FUNCTION_BLOCK FB_ActuatorModulating EXTENDS FB_Device
(*
	Continuous-position actuator: control valve, damper, any 0-100 % analog-positioned device.
	0 % = closed, 100 % = open. The output ramps to the setpoint at cfg.rampRate and is
	scaled to raw counts for an analog output terminal.
	
	Interlocks: losing them moves the actuator to cfg.safePosition. Permissives are required
	to move away from the safe position.
	
	Feedback: position comes from positionFdbk (FB_AnalogInput). In simulation, or with
	cfg.noFdbk, the position follows the output at the speed set by cfg.strokeTime.
	Simulation holds the physical output at 0.
*)
VAR_INPUT
	{attribute 'OPC.UA.DA' := '1'}
	{attribute 'OPC.UA.DA.StructuredType' := '1'}
	cfg					: ST_ActuatorModulatingConfiguration; //configuration
	
	{attribute 'OPC.UA.DA' := '1'}
	ocmd				: E_ActuatorModulatingCommand; //operator command
	{attribute 'OPC.UA.DA' := '1'}
	opPosition			: LREAL; //operator target position in %, used with ocmd Position
	
	func				: ST_ActuatorModulatingFunctions; //functions
	
	(* Interlocks/Permissives
	----------------------------------------------------------------------------------------------------*)
	{attribute 'OPC.UA.DA' := '1'}
	{attribute 'OPC.UA.DA.Access' := '1'}
	intlk				: FB_Permissive; //losing these moves the actuator to safePosition
	{attribute 'OPC.UA.DA' := '1'}
	{attribute 'OPC.UA.DA.Access' := '1'}
	perm				: FB_Permissive; //required to move away from safePosition
	
	(* External inputs
	----------------------------------------------------------------------------------------------------*)
	{attribute 'OPC.UA.DA' := '1'}
	{attribute 'OPC.UA.DA.Access' := '1'}
	positionFdbk		: FB_AnalogInput; //position feedback, link positionFdbk.inpRaw
END_VAR
VAR_OUTPUT
	outRaw		AT %Q*	: INT; //analog output to the actuator, link to the terminal's Value
	
	{attribute 'OPC.UA.DA' := '1'}
	{attribute 'OPC.UA.DA.Access' := '1'}
	{attribute 'OPC.UA.DA.StructuredType' := '1'}
	sts					: ST_ActuatorModulatingStatus;
	
	{attribute 'OPC.UA.DA' := '1'}
	{attribute 'OPC.UA.DA.Access' := '1'}
	{attribute 'OPC.UA.DA.StructuredType' := '1'}
	fault				: ST_ActuatorModulatingFault;
END_VAR
VAR
	//Command processing
	pcmd				: E_ActuatorModulatingCommand; //program command
	pPosition			: LREAL; //program target position in %, used with pcmd Position
	pcmdLast			: E_ActuatorModulatingCommand;
	ocmdLast			: E_ActuatorModulatingCommand;
	cmdReceived			: E_ActuatorModulatingCommand; //command accepted this scan
	targetReceived		: LREAL; //target position that came with cmdReceived
	funcTarget			: LREAL; //target of the running ToPosition function
	
	//state variables for tracking
	stateLastScan		: E_ActuatorModulatingState; //state on last scan
	simPosition			: LREAL; //simulated position in %
	
	//Oneshot triggers
	rtNewState			: BOOL; //just entered new state
	
	//Timers
	deltaTime			: FB_DeltaTime; //scan time for ramp and simulation
	positioningTimer	: TON; //time spent positioning
	
	resetFault			: BOOL;
END_VAR

SUPER^();

Device();
StatusIn();
ProcessInputs();
ProcessCommands();
Functions();
StateMachine();
HandleFaults();
ControlOutputs();
StatusOut();

METHOD PUBLIC Close
pcmd := E_ActuatorModulatingCommand.Close;
END_METHOD

METHOD PROTECTED ControlOutputs //Set physical outputs
IF sts.sim THEN //do not command outputs when simulated
	outRaw := 0;
ELSE
	outRaw := LREAL_TO_INT(F_ScaleLinear(value := sts.commandPosition, inMin := 0, inMax := 100,
										outMin := cfg.outRawAtClosed, outMax := cfg.outRawAtOpen, clamp := TRUE));
END_IF
END_METHOD

METHOD PROTECTED Device //map cfg to FB_Device and FB_Device to sts
// to FB device
opTimeout  			 := cfg.opTimeout;
opTimeoutEnable 	 := cfg.opTimeoutEnable;
opActivity 			 := ocmd <> E_ActuatorModulatingCommand.None;

// from FB device
sts.mode	   		 := mode;
sts.modeAuto   		 := sts.mode = E_SystemMode.Auto;
sts.modeManual 		 := sts.mode = E_SystemMode.Manual;
sts.manualOvrde		 := ctrl.manualOvrde;
sts.bypass 	   		 := ctrl.bypass;
sts.sim		   		 := ctrl.sim;
sts.parentConfigured := parentConfigured;
END_METHOD

METHOD PROTECTED Functions
VAR
	i : INT;
END_VAR
func.ToPosition(hmiTextStatic := CONCAT(cfg.actuatorId, ' to position'), timeoutPT := cfg.failTimePositioning);
func.ToPosition.permComplete.cfg.condText[0] := CONCAT(cfg.actuatorId, ' at position');
IF func.ToPosition.entry THEN
	funcTarget := sts.setpoint; // no Position parameter = stay where it is
	FOR i := GVL_Lib_SequencerConstants.MIN_PARAMETERS TO GVL_Lib_SequencerConstants.MAX_PARAMETERS DO
		IF func.ToPosition.arrParam[i].typeEnum = E_ActuatorModulatingFunctionParam.Position THEN
			funcTarget := func.ToPosition.arrParam[i].value;
		END_IF
	END_FOR
	SetPosition(funcTarget);
END_IF
IF func.ToPosition.running THEN
	func.ToPosition.permComplete.perm.0 := sts.atPosition AND ABS(sts.setpoint - LIMIT(cfg.minPosition, funcTarget, cfg.maxPosition)) < 0.001;
	IF NOT func.ToPosition.permComplete.perm.0 AND ABS(sts.setpoint - funcTarget) >= 0.001 AND NOT fault.active THEN
		SetPosition(funcTarget); // continue calling if didn't work at first
	END_IF
	func.ToPosition.inpError := fault.active;
	func.ToPosition.inpErrorText := fault.text;
END_IF


func.Open(hmiTextStatic := CONCAT(cfg.actuatorId, ' open'), timeoutPT := cfg.failTimePositioning);
func.Open.permComplete.cfg.condText[0] := CONCAT(cfg.actuatorId, ' open');
func.Open.permComplete.perm.0 := sts.atPosition AND sts.setpoint = cfg.maxPosition;
IF func.Open.entry OR (func.Open.running AND sts.setpoint <> cfg.maxPosition AND NOT fault.active) THEN
	Open();
END_IF
IF func.Open.running THEN
	func.Open.inpError := fault.active;
	func.Open.inpErrorText := fault.text;
END_IF


func.Close(hmiTextStatic := CONCAT(cfg.actuatorId, ' close'), timeoutPT := cfg.failTimePositioning);
func.Close.permComplete.cfg.condText[0] := CONCAT(cfg.actuatorId, ' closed');
func.Close.permComplete.perm.0 := sts.atPosition AND sts.setpoint = cfg.minPosition;
IF func.Close.entry OR (func.Close.running AND sts.setpoint <> cfg.minPosition AND NOT fault.active) THEN
	Close();
END_IF
IF func.Close.running THEN
	func.Close.inpError := fault.active;
	func.Close.inpErrorText := fault.text;
END_IF
END_METHOD

METHOD PROTECTED HandleFaults
fault.positionTimeout S= positioningTimer.Q;
fault.feedbackFault S= positionFdbk.fault.active AND NOT (cfg.noFdbk OR sts.sim);
//fault.intlkNOK; // Set in ProcessCommands and PrvPosition
//fault.permNOK; // Set in PrvPosition
//fault.ocmdNOK; // Set in ProcessCommands
//fault.pcmdNOK; // Set in ProcessCommands

(* ----- Handle Reset ----- *)
IF resetFault THEN
	fault.feedbackFault R= TRUE;
	fault.intlkNOK R= TRUE;
	fault.ocmdNOK R= TRUE;
	fault.pcmdNOK R= TRUE;
	fault.permNOK R= TRUE;
	fault.positionTimeout R= TRUE;
END_IF
resetFault := FALSE;

(* ----- Map Fault Id ----- *)
fault.id.0 := fault.feedbackFault;
fault.id.1 := fault.intlkNOK;
fault.id.2 := fault.ocmdNOK;
fault.id.3 := fault.pcmdNOK;
fault.id.4 := fault.permNOK;
fault.id.5 := fault.positionTimeout;

(* ----- Map Fault Text ----- *)
IF fault.feedbackFault THEN		fault.text := CONCAT(cfg.actuatorId, ' position feedback fault');
ELSIF fault.intlkNOK THEN		fault.text := CONCAT(cfg.actuatorId, ' interlocks not OK');
ELSIF fault.ocmdNOK THEN		fault.text := 'Operator command in Auto is not allowed';
ELSIF fault.pcmdNOK THEN		fault.text := 'Program command in Manual is not allowed';
ELSIF fault.permNOK THEN		fault.text := CONCAT(cfg.actuatorId, ' permissives not OK');
ELSIF fault.positionTimeout THEN	fault.text := CONCAT(cfg.actuatorId, ' did not reach position');
ELSE fault.text := '';
END_IF

(* ----- Set Active ----- *)
fault.active := fault.id > 0;
END_METHOD

METHOD PUBLIC Open
pcmd := E_ActuatorModulatingCommand.Open;
END_METHOD

METHOD PROTECTED ProcessCommands
//Check for new valid commands
IF ctrl.reset THEN
	PrvReset();
ELSIF ocmd <> E_ActuatorModulatingCommand.None THEN
	IF sts.modeManual THEN
		cmdReceived := ocmd;
		targetReceived := opPosition;
	ELSE
		fault.ocmdNOK := TRUE;
	END_IF
ELSIF pcmd <> E_ActuatorModulatingCommand.None THEN
	IF sts.modeAuto THEN
		cmdReceived := pcmd;
		targetReceived := pPosition;
	ELSE
		fault.pcmdNOK := TRUE;
	END_IF
END_IF

//Losing interlocks away from the safe position moves the actuator there
IF NOT intlk.sts.ok AND sts.setpoint <> cfg.safePosition THEN
	fault.intlkNOK S= TRUE;
	PrvSafe();
END_IF

CASE cmdReceived OF 
	E_ActuatorModulatingCommand.Close:
		PrvClose();
	E_ActuatorModulatingCommand.Open:
		PrvOpen();
	E_ActuatorModulatingCommand.Position:
		PrvPosition(targetReceived);
END_CASE

//Save last commands
IF pcmd <> E_ActuatorModulatingCommand.None THEN
	pcmdLast := pcmd;
END_IF
IF ocmd <> E_ActuatorModulatingCommand.None THEN
	ocmdLast := ocmd;
END_IF

//Clear commands every scan
cmdReceived	:= E_ActuatorModulatingCommand.None;
pcmd		:= E_ActuatorModulatingCommand.None;
ocmd		:= E_ActuatorModulatingCommand.None;
ctrl.reset	:= FALSE;
END_METHOD

METHOD PROTECTED ProcessInputs
deltaTime();

//Call input FBs
positionFdbk(cfg := cfg.positionFdbk);

//Use the simulated position when simulated or without feedback. Otherwise the simulated
//position tracks the real one, so switching to simulation does not jump.
IF cfg.noFdbk OR sts.sim THEN
	IF cfg.strokeTime > T#0S THEN
		simPosition := simPosition + LIMIT(-100.0 * deltaTime.seconds / (TIME_TO_LREAL(cfg.strokeTime) / 1000.0),
										   sts.commandPosition - simPosition,
										   100.0 * deltaTime.seconds / (TIME_TO_LREAL(cfg.strokeTime) / 1000.0));
	ELSE
		simPosition := sts.commandPosition;
	END_IF
	sts.position := simPosition;
ELSE
	sts.position := positionFdbk.sts.value;
	simPosition := sts.position;
END_IF
END_METHOD

METHOD PROTECTED PrvPosition
VAR_INPUT
	target		: LREAL; //requested position in %
END_VAR
VAR
	limited		: LREAL; //target within minPosition..maxPosition
END_VAR
limited := LIMIT(cfg.minPosition, target, cfg.maxPosition);

IF limited = sts.setpoint AND NOT sts.positioning THEN // ignore command if already there
	RETURN;
END_IF

IF limited = cfg.safePosition THEN // going to the safe position is always allowed
	PrvMove(limited);
ELSIF NOT intlk.sts.ok THEN // check intlk before moving away from safe
	fault.intlkNOK S= TRUE;
ELSIF NOT perm.sts.ok AND sts.setpoint = cfg.safePosition THEN // perm only needed to leave the safe position
	fault.permNOK S= TRUE;
ELSE
	PrvMove(limited);
END_IF
END_METHOD

METHOD PROTECTED PrvReset //Reset the device
resetFault S= TRUE;

//Reset permissives/interlocks and feedback
intlk.Reset();
perm.Reset();
positionFdbk.Reset();
END_METHOD

METHOD PROTECTED PrvSafe
sts.setpoint := cfg.safePosition;
sts.state := E_ActuatorModulatingState.Positioning;
END_METHOD

METHOD PUBLIC SetPosition
VAR_INPUT
	position	: LREAL; //target position in %
END_VAR
pPosition := position;
pcmd := E_ActuatorModulatingCommand.Position;
END_METHOD

METHOD PROTECTED StateMachine
//Ramp the output toward the setpoint
IF cfg.rampRate > 0 THEN
	sts.commandPosition := sts.commandPosition + LIMIT(-cfg.rampRate * deltaTime.seconds,
													   sts.setpoint - sts.commandPosition,
													   cfg.rampRate * deltaTime.seconds);
ELSE
	sts.commandPosition := sts.setpoint;
END_IF

sts.positionError := sts.setpoint - sts.position;

CASE sts.state OF
	
	E_ActuatorModulatingState.Positioning: //Check if we reached the setpoint
		IF ABS(sts.positionError) <= cfg.positionTolerance AND sts.commandPosition = sts.setpoint THEN
			sts.state := SettledState();
			sts.timeToPosition := positioningTimer.ET;
		END_IF
		
	E_ActuatorModulatingState.Closed,
	E_ActuatorModulatingState.Open,
	E_ActuatorModulatingState.AtPosition:
		// If we got here based on a successful move (which is the only way to get here), reset faults
		IF rtNewState THEN
			resetFault := TRUE;
		END_IF
		// Drifted off the setpoint: correct it
		IF ABS(sts.positionError) > MAX(cfg.driftTolerance, cfg.positionTolerance) THEN
			sts.state := E_ActuatorModulatingState.Positioning;
		ELSE
			sts.state := SettledState();
		END_IF
		
END_CASE

rtNewState := sts.state <> stateLastScan;
stateLastScan := sts.state;

// Monitoring timers
positioningTimer(IN := sts.state = E_ActuatorModulatingState.Positioning, PT := cfg.failTimePositioning);
END_METHOD

METHOD PROTECTED StatusIn
//Permissives and Interlocks
intlk(bypActive := sts.bypass, cfg := cfg.intlk);
perm(bypActive := sts.bypass, cfg := cfg.perm);
END_METHOD

METHOD PROTECTED StatusOut //Set output status information
sts.closed 		:= sts.state = E_ActuatorModulatingState.Closed;
sts.open 		:= sts.state = E_ActuatorModulatingState.Open;
sts.positioning	:= sts.state = E_ActuatorModulatingState.Positioning;
sts.atPosition	:= NOT sts.positioning;

sts.readyToMove	:= intlk.sts.ok AND perm.sts.ok;
sts.safe		:= NOT intlk.sts.ok AND sts.setpoint = cfg.safePosition;
sts.echoOutRaw	:= outRaw;
END_METHOD

METHOD PROTECTED PrvClose
PrvPosition(cfg.minPosition);
END_METHOD

METHOD PROTECTED PrvOpen
PrvPosition(cfg.maxPosition);
END_METHOD

METHOD PROTECTED SettledState : E_ActuatorModulatingState //state when at the setpoint
IF sts.position <= cfg.closedLimit THEN
	SettledState := E_ActuatorModulatingState.Closed;
ELSIF sts.position >= cfg.openLimit THEN
	SettledState := E_ActuatorModulatingState.Open;
ELSE
	SettledState := E_ActuatorModulatingState.AtPosition;
END_IF
END_METHOD

METHOD PROTECTED PrvMove //accept a new setpoint
VAR_INPUT
	target		: LREAL; //checked target position in %
END_VAR
sts.setpoint := target;
//Small trims (e.g. from a PID) stay settled; StateMachine starts positioning if the
//actuator falls behind by more than driftTolerance
IF ABS(target - sts.position) > cfg.positionTolerance THEN
	sts.state := E_ActuatorModulatingState.Positioning;
END_IF
END_METHOD

END_FUNCTION_BLOCK

(* stored: Version 1.1.0.1, ProductVersion 3.1.4024.12
   POU FB_ActuatorModulating: Id {43507db8-010e-47b6-b5b4-a9b43a020762}, SpecialFunc None
   Folder Protected: Id {0855584f-eb31-484c-a9db-066815d1c320}
   Folder Commands: Id {2c5a4f3c-27fe-4985-b773-17fc81068d3c}
   Folder Logic: Id {31c0ab04-64de-4302-a17e-6b26b2e5d911}
   Folder Public: Id {f0711d00-e70e-47ef-aeb3-0bd7d98dbc27}
   Folder Commands: Id {1ca77ccb-81b4-4c02-8673-f908cf8130ad}
   Method Close: Id {7457a5e1-323b-4c95-bd9b-940ce4e85636}
   Method ControlOutputs: Id {b8e8a569-0e3a-4b23-b043-4cf62bea2298}
   Method Device: Id {3092cebe-13b6-47f2-8c55-5d92fe2a9813}
   Method Functions: Id {9f0fabeb-8524-4bed-81d9-5743a0094e09}
   Method HandleFaults: Id {3c664065-467f-45bf-af80-27a24b791d17}
   Method Open: Id {53938b8c-a9be-4c81-8566-1bb197c18216}
   Method ProcessCommands: Id {a399af32-69a4-4773-8982-ea184bef2a85}
   Method ProcessInputs: Id {b1df521e-83fe-40ba-b7d8-2ff3f0869409}
   Method PrvPosition: Id {03aadde7-1384-4b87-aa0e-406e6569a9da}
   Method PrvReset: Id {b8966cc4-8c63-4b40-a6ac-aa5d2e75aab0}
   Method PrvSafe: Id {0a882f88-4765-4522-af42-64236a98b373}
   Method SetPosition: Id {73824b49-af45-4633-9006-8801b339ddde}
   Method StateMachine: Id {00cc7950-6830-4a7e-b9f1-91197a22503b}
   Method StatusIn: Id {d85b3c4b-6b37-4585-a33f-a44fe3de32c8}
   Method StatusOut: Id {2af30c99-9d64-4d2a-a8a7-a5d847c8a7ea}
   Method PrvClose: Id {7f775c9b-d081-44a6-82c5-4ae4f2441703}
   Method PrvOpen: Id {0fdbb7a4-f39e-4fc7-84bb-7a7ff0726101}
   Method SettledState: Id {6cb47ca7-dd0f-4127-a7a5-fba4293f3b3e}
   Method PrvMove: Id {c02d1281-c9dd-4fa5-a2d0-af0827d3bc6a} *)
